Fanuc KAREL source: kb00042.KL

PROGRAM KB00042
%STACKSIZE=65535
%PRIORITY=65535
%NOLOCKGROUP
VAR
P1 : STRING[80]
P2 : INTEGER
BEGIN
P1='A'
P2=1
CNV_STR_TIME(P1,P2)
END KB00042
